(* IEC 61131-3 sources: matiec/tests/var_list, 2 files *)

(* ---- decl_list.st ---- *)
TYPE PAIR : STRUCT
  A : UDINT;
  B : INT;
END_STRUCT; END_TYPE

FUNCTION_BLOCK FB1
  VAR
    T1, T2, T3 : TON;
  END_VAR
  T1(IN := TRUE, PT := T#1s);
END_FUNCTION_BLOCK

PROGRAM prog0
  VAR
    F : FB1;
    G1, G2, G3 : FB1;
    S1, S2, S3 : PAIR;
    N : INT;
  END_VAR
  F();
  N := N + 1;
END_PROGRAM

CONFIGURATION cfg
  RESOURCE res ON PLC
    TASK t(INTERVAL := T#10ms, PRIORITY := 0);
    PROGRAM inst WITH t : prog0;
  END_RESOURCE
END_CONFIGURATION

(* ---- struct_leaf.st ---- *)
TYPE INNER : STRUCT
  A : UDINT;
END_STRUCT; END_TYPE

TYPE OUTER : STRUCT
  X : UDINT;
  ARR : ARRAY[0..1] OF INT;
  S : STRING[7];
  IN1 : INNER;
END_STRUCT; END_TYPE

FUNCTION_BLOCK FB1
  VAR
    ST : OUTER;
  END_VAR
  ST.X := ST.X + 1;
END_FUNCTION_BLOCK

PROGRAM prog0
  VAR
    F : FB1;
    P : OUTER;
    N : INT;
  END_VAR
  F();
  N := N + 1;
END_PROGRAM

CONFIGURATION cfg
  RESOURCE res ON PLC
    TASK t(INTERVAL := T#10ms, PRIORITY := 0);
    PROGRAM inst WITH t : prog0;
  END_RESOURCE
END_CONFIGURATION
